FUNCTION_BLOCK Heating
VAR_INPUT
	diEnabled : BOOL;
	iSecImp : BOOL;
END_VAR
VAR_OUTPUT
	doEnabled : BOOL;
END_VAR
VAR_IN_OUT
	HeatingPhase : TPhaseHeating;
	Heater : THeater;
END_VAR
VAR
	pidParameters : ST_CTRL_PID_PARAMS;
END_VAR

{region "Aut/Man"}
    // switching state of engine - automatic or manual control (default state is manual)
    IF HeatingPhase.Cmd.AutCtrl AND NOT HeatingPhase.State.AutCtrl THEN
        HeatingPhase.State.AutCtrl := TRUE;
        HeatingPhase.State.ManCtrl := FALSE;
        HeatingPhase.State.Running := FALSE;
        HeatingPhase.State.Paused  := FALSE;
        HeatingPhase.State.Idle    := TRUE;
    ELSIF HeatingPhase.Cmd.ManCtrl AND NOT HeatingPhase.State.ManCtrl THEN
        HeatingPhase.State.ManCtrl := TRUE;
        HeatingPhase.State.AutCtrl := FALSE;
        HeatingPhase.State.Running := FALSE;
        HeatingPhase.State.Paused  := FALSE;
        HeatingPhase.State.Idle    := TRUE;
    END_IF;
    HeatingPhase.Cmd.AutCtrl := FALSE;
    HeatingPhase.Cmd.ManCtrl := FALSE;

    IF NOT HeatingPhase.State.AutCtrl AND NOT HeatingPhase.State.ManCtrl THEN
        HeatingPhase.State.ManCtrl := TRUE;
    END_IF;
{endregion}

{region "ManCtrl"}
    // processing manual actions - if command is processed, it is sets to FALSE even if can't be processed
    IF HeatingPhase.State.ManCtrl THEN
        // Start
        IF HeatingPhase.Cmd.StartMan AND HeatingPhase.State.Idle AND NOT Heater.State.GenErr THEN
            HeatingPhase.State.Idle    := FALSE;
            HeatingPhase.State.Running := TRUE;
            HeatingPhase.State.Done    := FALSE;
            Heater.Cmd.AutCtrl := TRUE;     // heater must be in auto, the phase drives it by request
        END_IF;

        // Pause
        IF HeatingPhase.Cmd.PauseMan AND HeatingPhase.State.Running THEN
            HeatingPhase.State.Running := FALSE;
            HeatingPhase.State.Paused  := TRUE;
        END_IF;

        // Resume
        IF HeatingPhase.Cmd.ResumeMan AND HeatingPhase.State.Paused AND NOT Heater.State.GenErr THEN
            HeatingPhase.State.Paused  := FALSE;
            HeatingPhase.State.Running := TRUE;
        END_IF;

        // Stop
        IF HeatingPhase.Cmd.StopMan AND (HeatingPhase.State.Running OR HeatingPhase.State.Paused) THEN
            HeatingPhase.State.Running := FALSE;
            HeatingPhase.State.Paused  := FALSE;
            HeatingPhase.State.Idle    := TRUE;
        END_IF;
    // real states of phase are writed into states in phase structure
    END_IF;

    HeatingPhase.Cmd.StartMan  := FALSE;
    HeatingPhase.Cmd.StopMan   := FALSE;
    HeatingPhase.Cmd.PauseMan  := FALSE;
    HeatingPhase.Cmd.ResumeMan := FALSE;
   
{endregion}

{region "AutCtrl"}
    // if request to run in automatic mode -> set auto request to heat to 1, if not request to heat 0
    // commands should be sets to false after their processing
    IF HeatingPhase.State.AutCtrl THEN
        IF HeatingPhase.Cmd.StartAut AND HeatingPhase.State.Idle AND NOT Heater.State.GenErr THEN
            HeatingPhase.State.Idle    := FALSE;
            HeatingPhase.State.Running := TRUE;
            HeatingPhase.State.Done    := FALSE;
            Heater.Cmd.AutCtrl := TRUE;
        END_IF;

        IF HeatingPhase.Cmd.StopAut AND (HeatingPhase.State.Running OR HeatingPhase.State.Paused) THEN
            HeatingPhase.State.Running := FALSE;
            HeatingPhase.State.Paused  := FALSE;
            HeatingPhase.State.Idle    := TRUE;
        END_IF;
    END_IF;

    HeatingPhase.Cmd.StartAut := FALSE;
    HeatingPhase.Cmd.StopAut  := FALSE;
{endregion}

{region "Done"}
    //every phase should have finish condition - heating phase - if water temp is on requested value for 10 seconds with 1°C hysteresis
    //after that done state should be setted to 1
    Heater.ThresholdTimer(
        IN := HeatingPhase.State.Running AND (ABS(HeatingPhase.WaterTemp - HeatingPhase.ParamReqTemp) <= 1.0),
        PT := T#10S);

    // time spent in the band, in seconds (for visualization)
    HeatingPhase.fTime := DINT_TO_INT(TIME_TO_DINT(Heater.ThresholdTimer.ET) / 1000);

    // finish condition
    IF HeatingPhase.State.Running AND Heater.ThresholdTimer.Q THEN
        HeatingPhase.State.Running := FALSE;
        HeatingPhase.State.Idle    := TRUE;
        HeatingPhase.State.Done    := TRUE;
    END_IF;

    // command reset done resets done state and than resets command
    IF HeatingPhase.Cmd.ResetDone THEN
        HeatingPhase.State.Done := FALSE;
        HeatingPhase.Cmd.ResetDone := FALSE;
    END_IF;
{endregion}

{region "States"}
    //Command valve in cases of states
    // Running - start heating  
    // Idle - stop heating
    // Pause - stop heating (alternative is hold actual temp)
    
    IF HeatingPhase.State.Running AND Heater.State.GenErr THEN
        HeatingPhase.State.Running := FALSE;
        HeatingPhase.State.Paused  := TRUE;
    END_IF;

    // setpoint for the PID controller in the heater
    Heater.ParamHeatingSetPointAutomat := HeatingPhase.ParamReqTemp;

    // Running - start heating
    // Idle    - stop heating
    // Paused  - stop heating (alternative would be to hold the actual temperature)
    Heater.Cmd.Req2RunAutCtrl := HeatingPhase.State.Running;
{endregion}

// delault state of phase - if not any state sets state to idle
IF NOT HeatingPhase.State.Idle AND NOT HeatingPhase.State.Paused AND NOT HeatingPhase.State.Running THEN
    HeatingPhase.State.Idle := 1;
END_IF;

doEnabled := diEnabled;

END_FUNCTION_BLOCK

(* stored: Version 1.1.0.1, ProductVersion 3.1.4024.13
   POU Heating: Id {67bfd793-3f9c-4f6b-ac3b-8ac7d5e1f5d7}, SpecialFunc None *)
